Staubli VAL3: DataBase4.dtx

public bool bAdjustXY_2_1
public bool bAdjustXY_2_2
public bool bAdjustXY_3_1
public bool bAdjustXY_3_2
public bool bAdjustXY_3_3
public bool bRefresh
public bool bShowJpos = true
public bool bTeach1 = true
public bool bTeach2 = true
public bool bTeach3
public bool bTeach4
public bool bTeach5
public bool bTeach6
public configRs cConfigSame
jointRs jA
public jointRs jAdjustXY_2_1 = {j1=26.957586, j2=-98.279005, j3=152.46178, j4=304.418255}
public jointRs jAdjustXY_2_2 = {j1=54.252313, j2=-89.434598, j3=152.46178, j4=88.28002}
public jointRs jAdjustXY_3_1
public jointRs jAdjustXY_3_2
public jointRs jAdjustXY_3_3
jointRs jB = {j4=365}
public jointRs jTeach1 = {j1=39.77131, j2=-98.855541, j3=9.53674E-05, j4=37.348709}
public jointRs jTeach2 = {j1=49.712231, j2=-94.333005, j3=-3.17891E-05, j4=-31.472397}
public jointRs jTeach3 = {j1=43.488119, j2=-71.195504, j3=-0.000127157, j4=-60.971375}
public jointRs jTeach4
public jointRs jTeach5
public jointRs jTeach6
public mdesc mSlow = {tmax=30, leave=0, reach=0, blend=cartesian}
public mdesc mSpeed_C_blend = {tmax=250, leave=0, reach=0, blend=cartesian}
public mdesc mSpeed_J_blend = {tmax=250, leave=5, reach=5}
public num nBtnItem = 82
public num nClock = 753.092
public num nJogMode
public num nStep0 = 21
public num nStep1 = 10
public num nStep2 = 10
public pointRs _pA = {x=519.21711, y=-79.50965, z=152.46178, rx=180, ry=5.610737E-15, rz=-143.096835, shoulder=lefty, fatherId=world[0]}
public pointRs _pB = {x=519.21711, y=-79.50965, z=152.46178, rx=180, ry=5.610737E-15, rz=-53.096835, shoulder=lefty, fatherId=world[0]}
public pointRs pAdjustXY_2_1 = {x=519.21711, y=-79.50965, z=152.46178, rx=180, ry=5.610737E-15, rz=126.903165, fatherId=world[0]}
public pointRs pAdjustXY_2_2 = {x=519.282115, y=-79.692376, z=152.46178, rx=-180, ry=-5.610803E-15, rz=-53.0977345, fatherId=world[0]}
public pointRs pAdjustXY_3_1 = {x=483.761349, y=-408.312989, z=81.104016, rx=180, ry=6.49774E-15, rz=112.169952, fatherId=world[0]}
public pointRs pAdjustXY_3_2 = {x=478.65297, y=-411.11562, z=81.104016, rx=180, ry=9.558925E-16, rz=172.169938, fatherId=world[0]}
public pointRs pAdjustXY_3_3 = {x=483.761365, y=-402.370049, z=81.104016, rx=-180, ry=5.541844E-15, rz=52.169883, fatherId=world[0]}
public pointRs pTeach1 = {x=507.856004, y=-117.232423, z=9.53674E-05, rx=-180, ry=2.598447E-15, rz=21.735523, shoulder=lefty, fatherId=world[0]}
public pointRs pTeach2 = {x=544.662238, y=-5.146269, z=-3.17891E-05, rx=-180, ry=6.811034E-15, rz=76.0931712, shoulder=lefty, fatherId=world[0]}
public pointRs pTeach3 = {x=647.536651, y=66.235993, z=-0.000127157, rx=-180, ry=7.014844E-15, rz=88.678759, fatherId=world[0]}
public pointRs pTeach4 = {x=384.117976, y=-405.930056, z=81.0572327, rx=180, ry=-7.012302E-15, rz=-91.97674, fatherId=world[0]}
public pointRs pTeach5 = {x=509.335923, y=-405.929869, z=81.0572327, rx=180, ry=-7.012305E-15, rz=-91.976094, fatherId=world[0]}
public pointRs pTeach6 = {x=509.281809, y=-464.347479, z=81.0572327, rx=180, ry=-7.012305E-15, rz=-91.976001, fatherId=world[0]}
string sAlertCN{}
  [Align] = "请按Move/Hold键对齐"
  [CantGoBack] = "不可重置!请首先记录第1点!"
  [CantMove1] = "不可到达!请重新记录第1点!"
  [CantMove2] = "不可到达!请重新记录这个点!"
  [CantSwitchTool2] = "不能切换tTool2!请先标定tTool1!"
  [CantSwitchTool3] = "不能切换tTool3!请先标定tTool2!"
  [CompleteAlign] = "对齐完成"
  [CompleteGoBack] = "重置完成"
  [CompleteMove] = "移动完成"
  [DeviationIsTooLarge] = "偏差过大!请重新记录点!"
  [Fifth] = "第5点记录完成"
  [First] = "第1点记录完成"
  [Fourth] = "第4点记录完成"
  [GoBack] = "请按Move/Hold键重置"
  [Move] = "请按Move/Hold键移动"
  [OffsetDone] = "偏差设置完成"
  [Quit] = "您是否决定退出TCP标定应用程序？"
  [SaveInTool1] = "工具参数保存在tTool1"
  [SaveInTool2] = "工具参数保存在tTool2"
  [SaveInTool3] = "工具参数保存在tTool3"
  [Second] = "第2点记录完成"
  [Seventh] = "第7点记录完成"
  [Sixth] = "第6点记录完成"
  [SwitchTool1] = "当前工具已经切换为tTool1!"
  [SwitchTool2] = "当前工具已经切换为tTool2!"
  [SwitchTool3] = "当前工具已经切换为tTool3!"
  [Third] = "第3点记录完成"
  [Version] = "版本: V2.1日期: 2020.10.12"
string sAlertEN{}
  [Align] = "Press Move/Hold Button To Align"
  [CantGoBack] = "Can't Go back!First record 1st point!"
  [CantMove1] = "Can't Reach!Re-record 1st point!"
  [CantMove2] = "Can't Reach!Re-record this point!"
  [CantSwitchTool2] = "Can't switch to tTool2!Please first calibrate tTool1!"
  [CantSwitchTool3] = "Can't switch to tTool3!Please first calibrate tTool2!"
  [CompleteAlign] = "Alignment has been completed"
  [CompleteGoBack] = "Go back has been completed"
  [CompleteMove] = "Movement has been completed"
  [DeviationIsTooLarge] = "Deviation is too large!Re-record points!"
  [Fifth] = "The 5th point has been recorded"
  [First] = "The 1st point has been recorded"
  [Fourth] = "The 4th point has been recorded"
  [GoBack] = "Press Move/Hold Button to Go back"
  [Move] = "Press Move/Hold Button to Move"
  [OffsetDone] = "Tool deviation has been enabled"
  [Quit] = "Are you sure to quit the tcp calibration application?"
  [SaveInTool1] = "Tool parameters are saved in tTool1"
  [SaveInTool2] = "Tool parameters are saved in tTool2"
  [SaveInTool3] = "Tool parameters are saved in tTool3"
  [Second] = "The 2nd point has been recorded"
  [Seventh] = "The 7th point has been recorded"
  [Sixth] = "The 6th point has been recorded"
  [SwitchTool1] = "The current tool has been switched to tTool1!"
  [SwitchTool2] = "The current tool has been switched to tTool2!"
  [SwitchTool3] = "The current tool has been switched to tTool3!"
  [Third] = "The 3rd point has been recorded"
  [Version] = "Version: V2.1 Date: October 12, 2020"
public string sCbxLanguage = "中文"
public string sCbxMounting = "置地"
string sHmiCN[200]
  [2] = "语言："
  [3] = "安装："
  [4] = "史陶比尔工具标定 - SmartTCP"
  [7] = "机型："
  [8] = "4轴"
  [9] = "6轴"
  [10] = "工具："
  [11] = "2点标定"
  [12] = "3点标定"
  [13] = "6点标定"
  [14] = "2点180°"
  [15] = "3点120°"
  [16] = "标定工具"
  [17] = "修正工具XY"
  [18] = "修正工具Z"
  [19] = "测试工具"
  [20] = "工具切换："
  [21] = "工具补偿："
  [31] = "点位：P1"
  [32] = "点位：P2"
  [33] = "点位：P3"
  [34] = "点位：P4"
  [35] = "点位：P5"
  [36] = "点位：P6"
  [41] = "步骤：1/2"
  [42] = "步骤：2/2"
  [43] = "步骤：1/3"
  [44] = "步骤：2/3"
  [45] = "步骤：3/3"
  [50] = "步骤：1/6"
  [51] = "步骤：2/6"
  [52] = "步骤：3/6"
  [53] = "步骤：4/6"
  [54] = "步骤：5/6"
  [55] = "步骤：6/6"
  [80] = "Null,记录,移动,Null,Null,Null,返回,继续"
  [81] = "Null,记录,移动,Null,Null,Null,返回,继续"
  [82] = "Null,记录,移动,Null,Null,计算,返回,完成"
  [83] = "Null,Null,Null,Null,Null,Null,Null,退出"
  [84] = "Null,记录,移动,切换,Null,Null,返回,继续"
  [85] = "重置,记录,移动,RZ+,RZ-,计算,返回,完成"
  [86] = "重置,记录,移动,RZ+,Null,Null,返回,继续"
  [87] = "重置,记录,移动,RZ-,Null,计算,返回,完成"
  [89] = "Null,Null,Null,Null,Null,Null,Null,完成"
  [100] = "适配TX2/TS2机器人的工具标定应用程序"
  [101] = "操作提醒："
  [102] = "工具垂直姿态对准尖点并记录"
  [103] = "工具任意姿态对准尖点并记录"
  [104] = "按计算按钮获取TCP值"
  [105] = "按记录按钮保存当前位置"
  [106] = "按记录按钮保存当前位置（坐标系原点）"
  [107] = "按记录按钮保存当前位置（坐标系OX方向）"
  [108] = "按记录按钮保存当前位置（坐标系OXY平面）"
  [109] = "保持当前姿态沿X方向移动"
  [110] = "保持当前姿态沿Y方向移动"
  [111] = "确保TCP(RZ) 可以反向旋转180°"
  [112] = "按RZ+(RZ-)与Move/Hold按钮旋转TCP 180°"
  [113] = "旋转TCP(RZ)接近一侧极限"
  [114] = "旋转TCP(RZ)接近中间位置"
  [115] = "确保TCP(RZ) 可以旋转±60°"
  [116] = "按RZ+与Move/Hold按钮旋转TCP +60°"
  [117] = "按RZ-与Move/Hold按钮旋转TCP -60°"
  [120] = "工具当前姿态对准尖点并记录"
  [121] = "最大可旋转角度只有:"
string sHmiEN[200]
  [2] = "Language："
  [3] = "Mounting："
  [4] = "Stäubli Tool Calibration - SmartTCP"
  [7] = "ArmType："
  [8] = "4axis"
  [9] = "6axis"
  [10] = "Tool："
  [11] = "2Points"
  [12] = "3Points"
  [13] = "6Points"
  [14] = "2Points180°"
  [15] = "3Points120°"
  [16] = "Calibration tool"
  [17] = "Correction tool XY"
  [18] = "Correction tool Z"
  [19] = "Verification tool"
  [20] = "Tool Switch："
  [21] = "Tool Offset："
  [31] = "Point：P1"
  [32] = "Point：P2"
  [33] = "Point：P3"
  [34] = "Point：P4"
  [35] = "Point：P5"
  [36] = "Point：P6"
  [41] = "Step：1/2"
  [42] = "Step：2/2"
  [43] = "Step：1/3"
  [44] = "Step：2/3"
  [45] = "Step：3/3"
  [50] = "Step：1/6"
  [51] = "Step：2/6"
  [52] = "Step：3/6"
  [53] = "Step：4/6"
  [54] = "Step：5/6"
  [55] = "Step：6/6"
  [80] = "Null,Here,Move,Null,Null,Null,Prev.,Next"
  [81] = "Null,Here,Move,Null,Null,Null,Prev.,Next"
  [82] = "Null,Here,Move,Null,Null,Calc.,Prev.,Done"
  [83] = "Null,Null,Null,Null,Null,Null,Null,Quit"
  [84] = "Null,Here,Move,Chg.,Null,Null,Prev.,Next"
  [85] = "Reset,Here,Move,RZ+,RZ-,Calc.,Prev.,Done"
  [86] = "Reset,Here,Move,RZ+,Null,Null,Prev.,Next"
  [87] = "Reset,Here,Move,RZ-,Null,Calc.,Prev.,Done"
  [89] = "Null,Null,Null,Null,Null,Null,Null,Done"
  [100] = "TCP calibration application for TX2/TS2 robot"
  [101] = "Operation reminder："
  [102] = "Touch to reference pointer in vertical attitude"
  [103] = "Touch to reference pointer in any attitude"
  [104] = "Press Calc. button to get the TCP value"
  [105] = "Press Here button to save the position"
  [106] = "Press Here button to save the position (Frame Origin)"
  [107] = "Press Here button to save the position (Frame Axis OX)"
  [108] = "Press Here button to save the position (Frame Plane OXY)"
  [109] = "Keep the current attitude moving in X direction"
  [110] = "Keep the current attitude moving in Y direction"
  [111] = "Ensure that the TCP(RZ) reverse can be rotated 180°"
  [112] = "Press the RZ+(RZ-) & Move/Hold to rotate TCP 180°"
  [113] = "Rotate TCP (RZ) close to one side limit"
  [114] = "Rotate TCP (RZ) close to middle position"
  [115] = "Ensure that the TCP(RZ) can be rotated ±60°"
  [116] = "Press the RZ+ & Move/Hold to rotate TCP +60°"
  [117] = "Press the RZ- & Move/Hold to rotate TCP -60°"
  [120] = "Touch to reference pointer in current attitude"
  [121] = "The maximum rotation angle is only:"
public string sLanguage = "chinese"
public string sLanguageM = "chinese"
public string sMounting = "Floor"
public tool tCurrentTool = {fatherId=flange[0]}
public tool tFlange = {fatherId=flange[0]}
public tool tTool1 = {x=119.999929, y=55.000162261, fatherId=flange[0], ioLink=FastIO\fOut0}
public tool tTool2 = {x=-144.465483, y=50.826546, fatherId=flange[0], ioLink=FastIO\fOut0}
public trsf trOffset = {z=10}
public trsf trOffsetM = {x=11, y=22, z=33, rx=44, ry=55, rz=66}
public utButton utBtn_Bottom[8]
  [0]
    utAppearance Appearance
      [0]
        bool bVisibility
        string sBackgroundColour = "#FFFFFF"
        string sBackgroundImage
        string sColour
    utBorder Border
      [0]
        string sBorderColour
    utCommon Common
      [0]
        bool bDisabled
        string sID = "bottom_btn0"
        string sPage = "Disk://SmartTCP_CS9/ts2/interface/Page_Main"
        string sText
    utData Data
      [0]
        bool bStatus
        num nVal
    utEvents Events
      [0]
        bool bClick
        bool bMouseDown
        bool bMouseUp
    utText Text
      [0]
        num nFontSize
        string sFontFamily
        string sFontStyle
        string sFontWeight
        string sTextAlignment
  [1]
    utAppearance Appearance
      [0]
        bool bVisibility = true
        string sBackgroundColour = "#FFFFFF"
        string sBackgroundImage
        string sColour
    utBorder Border
      [0]
        string sBorderColour
    utCommon Common
      [0]
        bool bDisabled
        string sID = "bottom_btn1"
        string sPage = "Disk://SmartTCP_CS9/ts2/interface/Page_Main"
        string sText = "记录"
    utData Data
      [0]
        bool bStatus
        num nVal
    utEvents Events
      [0]
        bool bClick
        bool bMouseDown
        bool bMouseUp
    utText Text
      [0]
        num nFontSize
        string sFontFamily
        string sFontStyle
        string sFontWeight
        string sTextAlignment
  [2]
    utAppearance Appearance
      [0]
        bool bVisibility = true
        string sBackgroundColour = "#FFFFFF"
        string sBackgroundImage
        string sColour
    utBorder Border
      [0]
        string sBorderColour
    utCommon Common
      [0]
        bool bDisabled
        string sID = "bottom_btn2"
        string sPage = "Disk://SmartTCP_CS9/ts2/interface/Page_Main"
        string sText = "移动"
    utData Data
      [0]
        bool bStatus
        num nVal
    utEvents Events
      [0]
        bool bClick
        bool bMouseDown
        bool bMouseUp
    utText Text
      [0]
        num nFontSize
        string sFontFamily
        string sFontStyle
        string sFontWeight
        string sTextAlignment
  [3]
    utAppearance Appearance
      [0]
        bool bVisibility
        string sBackgroundColour = "#FFFFFF"
        string sBackgroundImage
        string sColour
    utBorder Border
      [0]
        string sBorderColour
    utCommon Common
      [0]
        bool bDisabled
        string sID = "bottom_btn3"
        string sPage = "Disk://SmartTCP_CS9/ts2/interface/Page_Main"
        string sText
    utData Data
      [0]
        bool bStatus
        num nVal
    utEvents Events
      [0]
        bool bClick
        bool bMouseDown
        bool bMouseUp
    utText Text
      [0]
        num nFontSize
        string sFontFamily
        string sFontStyle
        string sFontWeight
        string sTextAlignment
  [4]
    utAppearance Appearance
      [0]
        bool bVisibility
        string sBackgroundColour = "#FFFFFF"
        string sBackgroundImage
        string sColour
    utBorder Border
      [0]
        string sBorderColour
    utCommon Common
      [0]
        bool bDisabled
        string sID = "bottom_btn4"
        string sPage = "Disk://SmartTCP_CS9/ts2/interface/Page_Main"
        string sText
    utData Data
      [0]
        bool bStatus
        num nVal
    utEvents Events
      [0]
        bool bClick
        bool bMouseDown
        bool bMouseUp
    utText Text
      [0]
        num nFontSize
        string sFontFamily
        string sFontStyle
        string sFontWeight
        string sTextAlignment
  [5]
    utAppearance Appearance
      [0]
        bool bVisibility = true
        string sBackgroundColour = "#FFFFFF"
        string sBackgroundImage
        string sColour
    utBorder Border
      [0]
        string sBorderColour
    utCommon Common
      [0]
        bool bDisabled
        string sID = "bottom_btn5"
        string sPage = "Disk://SmartTCP_CS9/ts2/interface/Page_Main"
        string sText = "计算"
    utData Data
      [0]
        bool bStatus
        num nVal
    utEvents Events
      [0]
        bool bClick
        bool bMouseDown
        bool bMouseUp
    utText Text
      [0]
        num nFontSize
        string sFontFamily
        string sFontStyle
        string sFontWeight
        string sTextAlignment
  [6]
    utAppearance Appearance
      [0]
        bool bVisibility = true
        string sBackgroundColour = "#FFFFFF"
        string sBackgroundImage
        string sColour
    utBorder Border
      [0]
        string sBorderColour
    utCommon Common
      [0]
        bool bDisabled
        string sID = "bottom_btn6"
        string sPage = "Disk://SmartTCP_CS9/ts2/interface/Page_Main"
        string sText = "返回"
    utData Data
      [0]
        bool bStatus
        num nVal
    utEvents Events
      [0]
        bool bClick
        bool bMouseDown
        bool bMouseUp
    utText Text
      [0]
        num nFontSize
        string sFontFamily
        string sFontStyle
        string sFontWeight
        string sTextAlignment
  [7]
    utAppearance Appearance
      [0]
        bool bVisibility = true
        string sBackgroundColour = "#FFFFFF"
        string sBackgroundImage
        string sColour
    utBorder Border
      [0]
        string sBorderColour
    utCommon Common
      [0]
        bool bDisabled
        string sID = "bottom_btn7"
        string sPage = "Disk://SmartTCP_CS9/ts2/interface/Page_Main"
        string sText = "完成"
    utData Data
      [0]
        bool bStatus
        num nVal
    utEvents Events
      [0]
        bool bClick
        bool bMouseDown
        bool bMouseUp
    utText Text
      [0]
        num nFontSize
        string sFontFamily
        string sFontStyle
        string sFontWeight
        string sTextAlignment
public utButton utBtn_No
  [0]
    utAppearance Appearance
      [0]
        bool bVisibility = true
        string sBackgroundColour = "#FFFFFF"
        string sBackgroundImage
        string sColour
    utBorder Border
      [0]
        string sBorderColour
    utCommon Common
      [0]
        bool bDisabled
        string sID = "btn_No"
        string sPage = "Disk://SmartTCP_CS9/ts2/interface/Page_Container_Confirm"
        string sText = "No"
    utData Data
      [0]
        bool bStatus
        num nVal
    utEvents Events
      [0]
        bool bClick
        bool bMouseDown
        bool bMouseUp
    utText Text
      [0]
        num nFontSize
        string sFontFamily
        string sFontStyle
        string sFontWeight
        string sTextAlignment
public utButton utBtn_OK
  [0]
    utAppearance Appearance
      [0]
        bool bVisibility = true
        string sBackgroundColour = "#FFFFFF"
        string sBackgroundImage
        string sColour
    utBorder Border
      [0]
        string sBorderColour
    utCommon Common
      [0]
        bool bDisabled
        string sID = "btn_OK"
        string sPage = "Disk://SmartTCP_CS9/ts2/interface/Page_Container_Alert"
        string sText = "OK"
    utData Data
      [0]
        bool bStatus
        num nVal
    utEvents Events
      [0]
        bool bClick
        bool bMouseDown
        bool bMouseUp
    utText Text
      [0]
        num nFontSize
        string sFontFamily
        string sFontStyle
        string sFontWeight
        string sTextAlignment
public utButton utBtn_Step[3]
  [0]
    utAppearance Appearance
      [0]
        bool bVisibility = true
        string sBackgroundColour = "#FFFFFF"
        string sBackgroundImage
        string sColour
    utBorder Border
      [0]
        string sBorderColour
    utCommon Common
      [0]
        bool bDisabled
        string sID = "step_btn0"
        string sPage = "Disk://SmartTCP_CS9/ts2/interface/Page_Container_Main"
        string sText = "标定工具"
    utData Data
      [0]
        bool bStatus
        num nVal = 16
    utEvents Events
      [0]
        bool bClick = true
        bool bMouseDown
        bool bMouseUp
    utText Text
      [0]
        num nFontSize
        string sFontFamily
        string sFontStyle
        string sFontWeight
        string sTextAlignment
  [1]
    utAppearance Appearance
      [0]
        bool bVisibility = true
        string sBackgroundColour = "#FFFFFF"
        string sBackgroundImage
        string sColour
    utBorder Border
      [0]
        string sBorderColour
    utCommon Common
      [0]
        bool bDisabled
        string sID = "step_btn1"
        string sPage = "Disk://SmartTCP_CS9/ts2/interface/Page_Container_Main"
        string sText = "修正工具XY"
    utData Data
      [0]
        bool bStatus
        num nVal = 17
    utEvents Events
      [0]
        bool bClick
        bool bMouseDown
        bool bMouseUp
    utText Text
      [0]
        num nFontSize
        string sFontFamily
        string sFontStyle
        string sFontWeight
        string sTextAlignment
  [2]
    utAppearance Appearance
      [0]
        bool bVisibility = true
        string sBackgroundColour = "#FFFFFF"
        string sBackgroundImage
        string sColour
    utBorder Border
      [0]
        string sBorderColour
    utCommon Common
      [0]
        bool bDisabled
        string sID = "step_btn2"
        string sPage = "Disk://SmartTCP_CS9/ts2/interface/Page_Container_Main"
        string sText = "测试工具"
    utData Data
      [0]
        bool bStatus
        num nVal = 19
    utEvents Events
      [0]
        bool bClick
        bool bMouseDown
        bool bMouseUp
    utText Text
      [0]
        num nFontSize
        string sFontFamily
        string sFontStyle
        string sFontWeight
        string sTextAlignment
public utButton utBtn_Yes
  [0]
    utAppearance Appearance
      [0]
        bool bVisibility = true
        string sBackgroundColour = "#FFFFFF"
        string sBackgroundImage
        string sColour
    utBorder Border
      [0]
        string sBorderColour
    utCommon Common
      [0]
        bool bDisabled
        string sID = "btn_Yes"
        string sPage = "Disk://SmartTCP_CS9/ts2/interface/Page_Container_Confirm"
        string sText = "Yes"
    utData Data
      [0]
        bool bStatus
        num nVal
    utEvents Events
      [0]
        bool bClick
        bool bMouseDown
        bool bMouseUp
    utText Text
      [0]
        num nFontSize
        string sFontFamily
        string sFontStyle
        string sFontWeight
        string sTextAlignment
public utCombo utCbx_Language_Data
  [0]
    utAppearance Appearance
      [0]
        bool bVisibility
        string sBackgroundColour
        string sColour
    utBorder Border
      [0]
        string sBorderColour
        string sBorderStyle
        string sBorderWidth
    utCommon Common
      [0]
        bool bDisabled
        string sID = "cbx_Language_D"
        string sItem[2]
          [0] = "中文"
          [1] = "英文"
        string sOption{}
        string sPage = "Disk://SmartTCP_CS9/ts2/interface/Page_Main"
        string sValue = "中文"
    utData Data
      [0]
        bool bStatus
        num nVal
    utText Text
      [0]
        num nFontSize
        string sFontFamily
        string sFontStyle
public utCombo utCbx_Mounting_Data
  [0]
    utAppearance Appearance
      [0]
        bool bVisibility
        string sBackgroundColour
        string sColour
    utBorder Border
      [0]
        string sBorderColour
        string sBorderStyle
        string sBorderWidth
    utCommon Common
      [0]
        bool bDisabled
        string sID = "cbx_Mounting_D"
        string sItem[2]
          [0] = "置地"
          [1] = "置顶"
        string sOption{}
        string sPage = "Disk://SmartTCP_CS9/ts2/interface/Page_Main"
        string sValue = "置地"
    utData Data
      [0]
        bool bStatus
        num nVal
    utText Text
      [0]
        num nFontSize
        string sFontFamily
        string sFontStyle
public utContainer utCtn_Function
  [0]
    utAppearance Appearance
      [0]
        bool bVisibility = true
    utCommon Common
      [0]
        string sID = "ctn_Function"
        string sPage = "Disk://SmartTCP_CS9/ts2/interface/Page_Main"
        string sSource = "Page_Container_Teach.html"
public utContainer utCtn_Message
  [0]
    utAppearance Appearance
      [0]
        bool bVisibility = true
    utCommon Common
      [0]
        string sID = "ctn_Message"
        string sPage = "Disk://SmartTCP_CS9/ts2/interface/Page_Main"
        string sSource = "Page_Container_Alert.html"
public utImage utImg_CheckBox_a[3]
  [0]
    utAppearance Appearance
      [0]
        bool bVisibility
        string sBackgroundColour
    utBorder Border
      [0]
        num nBorderWidth
        string sBorderColour
        string sBorderStyle
    utCommon Common
      [0]
        string sClass = "clickable"
        string sID = "img_CheckBox_a0"
        string sPage = "Disk://SmartTCP_CS9/ts2/interface/Page_Container_Main"
        string sSourceImage = "images/checkbox_checked.png"
    utData Data
      [0]
        bool bStatus = true
        num nVal
        string sSourceImg1 = "images/checkbox_checked.png"
        string sSourceImg2 = "images/checkbox_unchecked.png"
    utEvents Events
      [0]
        bool bClick
        bool bMouseDown
        bool bMouseUp
  [1]
    utAppearance Appearance
      [0]
        bool bVisibility
        string sBackgroundColour
    utBorder Border
      [0]
        num nBorderWidth
        string sBorderColour
        string sBorderStyle
    utCommon Common
      [0]
        string sClass = "clickable"
        string sID = "img_CheckBox_a1"
        string sPage = "Disk://SmartTCP_CS9/ts2/interface/Page_Container_Main"
        string sSourceImage = "images/checkbox_unchecked.png"
    utData Data
      [0]
        bool bStatus
        num nVal
        string sSourceImg1 = "images/checkbox_checked.png"
        string sSourceImg2 = "images/checkbox_unchecked.png"
    utEvents Events
      [0]
        bool bClick
        bool bMouseDown
        bool bMouseUp
  [2]
    utAppearance Appearance
      [0]
        bool bVisibility
        string sBackgroundColour
    utBorder Border
      [0]
        num nBorderWidth
        string sBorderColour
        string sBorderStyle
    utCommon Common
      [0]
        string sClass = "clickable"
        string sID = "img_CheckBox_a2"
        string sPage = "Disk://SmartTCP_CS9/ts2/interface/Page_Container_Main"
        string sSourceImage = "images/checkbox_unchecked.png"
    utData Data
      [0]
        bool bStatus
        num nVal
        string sSourceImg1 = "images/checkbox_checked.png"
        string sSourceImg2 = "images/checkbox_unchecked.png"
    utEvents Events
      [0]
        bool bClick
        bool bMouseDown
        bool bMouseUp
public utImage utImg_CheckBox_b[2]
  [0]
    utAppearance Appearance
      [0]
        bool bVisibility
        string sBackgroundColour
    utBorder Border
      [0]
        num nBorderWidth
        string sBorderColour
        string sBorderStyle
    utCommon Common
      [0]
        string sClass = "clickable"
        string sID = "img_CheckBox_b0"
        string sPage = "Disk://SmartTCP_CS9/ts2/interface/Page_Container_Main"
        string sSourceImage = "images/checkbox_checked.png"
    utData Data
      [0]
        bool bStatus = true
        num nVal
        string sSourceImg1 = "images/checkbox_checked.png"
        string sSourceImg2 = "images/checkbox_unchecked.png"
    utEvents Events
      [0]
        bool bClick
        bool bMouseDown
        bool bMouseUp
  [1]
    utAppearance Appearance
      [0]
        bool bVisibility
        string sBackgroundColour
    utBorder Border
      [0]
        num nBorderWidth
        string sBorderColour
        string sBorderStyle
    utCommon Common
      [0]
        string sClass = "clickable"
        string sID = "img_CheckBox_b1"
        string sPage = "Disk://SmartTCP_CS9/ts2/interface/Page_Container_Main"
        string sSourceImage = "images/checkbox_unchecked.png"
    utData Data
      [0]
        bool bStatus
        num nVal
        string sSourceImg1 = "images/checkbox_checked.png"
        string sSourceImg2 = "images/checkbox_unchecked.png"
    utEvents Events
      [0]
        bool bClick
        bool bMouseDown
        bool bMouseUp
public utImage utImg_Example
  [0]
    utAppearance Appearance
      [0]
        bool bVisibility = true
        string sBackgroundColour
    utBorder Border
      [0]
        num nBorderWidth
        string sBorderColour
        string sBorderStyle
    utCommon Common
      [0]
        string sClass = "clickable"
        string sID = "img_example"
        string sPage = "Disk://SmartTCP_CS9/ts2/interface/Page_Container_Teach"
        string sSourceImage = "images/4AxisTeach_2.jpg"
    utData Data
      [0]
        bool bStatus
        num nVal
        string sSourceImg1
        string sSourceImg2
    utEvents Events
      [0]
        bool bClick
        bool bMouseDown
        bool bMouseUp
public utImage utImg_Info
  [0]
    utAppearance Appearance
      [0]
        bool bVisibility = true
        string sBackgroundColour
    utBorder Border
      [0]
        num nBorderWidth
        string sBorderColour
        string sBorderStyle
    utCommon Common
      [0]
        string sClass = "clickable"
        string sID = "img_info"
        string sPage = "Disk://SmartTCP_CS9/ts2/interface/Page_Main"
        string sSourceImage = "images/info.png"
    utData Data
      [0]
        bool bStatus
        num nVal
        string sSourceImg1 = "images/switch_on.png"
        string sSourceImg2 = "images/switch_off.png"
    utEvents Events
      [0]
        bool bClick
        bool bMouseDown
        bool bMouseUp
public utImage utImg_JogMode[4]
  [0]
    utAppearance Appearance
      [0]
        bool bVisibility = true
        string sBackgroundColour
    utBorder Border
      [0]
        num nBorderWidth
        string sBorderColour = "#FFFFFF"
        string sBorderStyle = "None"
    utCommon Common
      [0]
        string sClass = "selected"
        string sID = "img_None"
        string sPage = "Disk://SmartTCP_CS9/ts2/interface/Page_Main"
        string sSourceImage = "images/none.svg"
    utData Data
      [0]
        bool bStatus
        num nVal
        string sSourceImg1
        string sSourceImg2
    utEvents Events
      [0]
        bool bClick
        bool bMouseDown
        bool bMouseUp
  [1]
    utAppearance Appearance
      [0]
        bool bVisibility = true
        string sBackgroundColour
    utBorder Border
      [0]
        num nBorderWidth
        string sBorderColour = "#FFFFFF"
        string sBorderStyle = "None"
    utCommon Common
      [0]
        string sClass = "clickable"
        string sID = "img_Joint"
        string sPage = "Disk://SmartTCP_CS9/ts2/interface/Page_Main"
        string sSourceImage = "images/joint.svg"
    utData Data
      [0]
        bool bStatus
        num nVal
        string sSourceImg1
        string sSourceImg2
    utEvents Events
      [0]
        bool bClick
        bool bMouseDown
        bool bMouseUp
  [2]
    utAppearance Appearance
      [0]
        bool bVisibility = true
        string sBackgroundColour
    utBorder Border
      [0]
        num nBorderWidth
        string sBorderColour = "#000000"
        string sBorderStyle = "Solid"
    utCommon Common
      [0]
        string sClass = "clickable"
        string sID = "img_Frame"
        string sPage = "Disk://SmartTCP_CS9/ts2/interface/Page_Main"
        string sSourceImage = "images/frame.svg"
    utData Data
      [0]
        bool bStatus
        num nVal
        string sSourceImg1
        string sSourceImg2
    utEvents Events
      [0]
        bool bClick
        bool bMouseDown
        bool bMouseUp
  [3]
    utAppearance Appearance
      [0]
        bool bVisibility = true
        string sBackgroundColour
    utBorder Border
      [0]
        num nBorderWidth
        string sBorderColour = "#FFFFFF"
        string sBorderStyle = "None"
    utCommon Common
      [0]
        string sClass = "clickable"
        string sID = "img_Tool"
        string sPage = "Disk://SmartTCP_CS9/ts2/interface/Page_Main"
        string sSourceImage = "images/tool.svg"
    utData Data
      [0]
        bool bStatus
        num nVal
        string sSourceImg1
        string sSourceImg2
    utEvents Events
      [0]
        bool bClick
        bool bMouseDown
        bool bMouseUp
public utImage utImg_Next
  [0]
    utAppearance Appearance
      [0]
        bool bVisibility = true
        string sBackgroundColour
    utBorder Border
      [0]
        num nBorderWidth
        string sBorderColour
        string sBorderStyle
    utCommon Common
      [0]
        string sClass = "clickable"
        string sID = "img_Next"
        string sPage = "Disk://SmartTCP_CS9/ts2/interface/Page_Container_Test"
        string sSourceImage = "images/navigate-next.svg"
    utData Data
      [0]
        bool bStatus
        num nVal
        string sSourceImg1
        string sSourceImg2
    utEvents Events
      [0]
        bool bClick
        bool bMouseDown
        bool bMouseUp
public utImage utImg_PosSwitch
  [0]
    utAppearance Appearance
      [0]
        bool bVisibility = true
        string sBackgroundColour
    utBorder Border
      [0]
        num nBorderWidth
        string sBorderColour
        string sBorderStyle
    utCommon Common
      [0]
        string sClass = "clickable"
        string sID = "img_PosSwitch"
        string sPage = "Disk://SmartTCP_CS9/ts2/interface/Page_Main"
        string sSourceImage = "images/switch.png"
    utData Data
      [0]
        bool bStatus
        num nVal
        string sSourceImg1
        string sSourceImg2
    utEvents Events
      [0]
        bool bClick
        bool bMouseDown
        bool bMouseUp
public utImage utImg_Previous
  [0]
    utAppearance Appearance
      [0]
        bool bVisibility = true
        string sBackgroundColour
    utBorder Border
      [0]
        num nBorderWidth
        string sBorderColour
        string sBorderStyle
    utCommon Common
      [0]
        string sClass = "clickable"
        string sID = "img_Previous"
        string sPage = "Disk://SmartTCP_CS9/ts2/interface/Page_Container_Test"
        string sSourceImage = "images/navigate-previous.svg"
    utData Data
      [0]
        bool bStatus
        num nVal
        string sSourceImg1
        string sSourceImg2
    utEvents Events
      [0]
        bool bClick
        bool bMouseDown
        bool bMouseUp
public utImage utImg_Switch
  [0]
    utAppearance Appearance
      [0]
        bool bVisibility
        string sBackgroundColour
    utBorder Border
      [0]
        num nBorderWidth
        string sBorderColour
        string sBorderStyle
    utCommon Common
      [0]
        string sClass = "clickable"
        string sID = "img_Switch"
        string sPage = "Disk://SmartTCP_CS9/ts2/interface/Page_Container_Test"
        string sSourceImage = "images/switch_off.png"
    utData Data
      [0]
        bool bStatus
        num nVal
        string sSourceImg1 = "images/switch_on.png"
        string sSourceImg2 = "images/switch_off.png"
    utEvents Events
      [0]
        bool bClick
        bool bMouseDown
        bool bMouseUp
public utLabel utLbl_Axis
  [0]
    utAppearance Appearance
      [0]
        bool bVisibility
        string sBackgroundColour = "#FFFFFF"
        string sColour
    utBorder Border
      [0]
        num nBorderWidth
        string sBorderColour
        string sBorderStyle
    utCommon Common
      [0]
        string sID = "lbl_Axis"
        string sPage = "Disk://SmartTCP_CS9/ts2/interface/Page_Main"
        string sText = "机型："
    utData Data
      [0]
        bool bStatus
        num nVal = 99
    utEvents Events
      [0]
        bool bClick
        bool bMouseDown
        bool bMouseUp
    utText Text
      [0]
        num nFontSize
        string sFontFamily
        string sFontStyle
        string sFontWeight
        string sTextAlignment
public utLabel utLbl_Axis_Data
  [0]
    utAppearance Appearance
      [0]
        bool bVisibility
        string sBackgroundColour = "#FFFFFF"
        string sColour
    utBorder Border
      [0]
        num nBorderWidth
        string sBorderColour
        string sBorderStyle
    utCommon Common
      [0]
        string sID = "lbl_Axis_Data"
        string sPage = "Disk://SmartTCP_CS9/ts2/interface/Page_Main"
        string sText = "4轴"
    utData Data
      [0]
        bool bStatus
        num nVal = 99
    utEvents Events
      [0]
        bool bClick
        bool bMouseDown
        bool bMouseUp
    utText Text
      [0]
        num nFontSize
        string sFontFamily
        string sFontStyle
        string sFontWeight
        string sTextAlignment
public utLabel utLbl_CheckBox_a[3]
  [0]
    utAppearance Appearance
      [0]
        bool bVisibility
        string sBackgroundColour = "#FFFFFF"
        string sColour
    utBorder Border
      [0]
        num nBorderWidth
        string sBorderColour
        string sBorderStyle
    utCommon Common
      [0]
        string sID = "lbl_CheckBox_a0"
        string sPage = "Disk://SmartTCP_CS9/ts2/interface/Page_Container_Main"
        string sText = "2点标定"
    utData Data
      [0]
        bool bStatus
        num nVal = 99
    utEvents Events
      [0]
        bool bClick
        bool bMouseDown
        bool bMouseUp
    utText Text
      [0]
